Fanuc KAREL source: KA00024.KL

PROGRAM KA00024
%NOLOCKGROUP
VAR
  SRC: REAL
  DST: ARRAY[2] OF SHORT
BEGIN
  SRC = 2.0
  DST[1] = SRC
END KA00024
